% RSLogix 500 project L12c_operation on analog ip op.RSS, saved by version 8.30.00.16 %
PROJECT "UNTITLED"    % processor: MicroLogix 1000 %

PROGRAM FILES
  LAD 2 "MAIN_PROG"  4 rungs
  LAD 3 "USER_FAULT"  1 rungs
  LAD 4 "HSC_INT"  1 rungs
  LAD 5 "STI_INT"  1 rungs
  LAD 6, 7, 8, 9, 10, 11, 12, 13, 14, 15, 16: only END

DATA FILES
  O0 OUTPUT  5 elements
  I1 INPUT  8 elements
  S2 STATUS  33 elements
  B3 BINARY  32 elements
  T4 TIMER  40 elements
  C5 COUNTER  32 elements
  R6 CONTROL  16 elements
  N7 INTEGER  105 elements

LADDER 2 "MAIN_PROG"
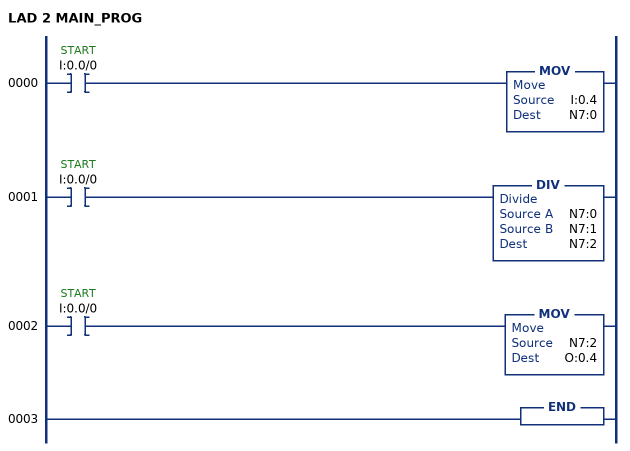
% Rung: 0 %
SOR XIC I:0.0/0 MOV I:0.4 N7:0 EOR
%   I:0.0/0  "START" %
%   I:0.4  "analog input 1 address" %
% Rung: 1 %
SOR XIC I:0.0/0 DIV N7:0 N7:1 N7:2 EOR
%   I:0.0/0  "START" %
% Rung: 2 %
SOR XIC I:0.0/0 MOV N7:2 O:0.4 EOR
%   I:0.0/0  "START" %
% Rung: 3 %
SOR END EOR

DATA TABLE (non-zero values as saved)
DATA N7
% N7:0 % 10 2 5 0 0 0 0 0 0 0
